	IF fbStopTx.bSettled THEN
		fbHourAngle.StopAxis := FALSE;
		fbDeclination.StopAxis := FALSE;
		_StopTelescope := FALSE;
	END_IF
END_IF
END_METHOD

METHOD PRIVATE _TrackTelescope : BOOL
VAR_INPUT
END_VAR
// send Dome position
THIS^.fbDome.Position := fAzimuthCurrent;
// Declination (including offest and pointing model)
fbDeclination.Position := fDeclinationApparent + fDeclinationOffset + fDeclinationPointingOffset;
// HourAngle
// change to -180 to 180 degree in HA
IF MODABS(fHourAngleApparent + F_HourAngleOffsetOnAxis(fHourAngleOffset, fDeclinationApparent)+ fHourAnglePointingOffset, 360) > 180 THEN
	fbHourAngle.Position := MODABS(fHourAngleApparent + F_HourAngleOffsetOnAxis(fHourAngleOffset, fDeclinationApparent)+ fHourAnglePointingOffset,360) - 360.0;
ELSE
	fbHourAngle.Position := MODABS(fHourAngleApparent + F_HourAngleOffsetOnAxis(fHourAngleOffset, fDeclinationApparent)+ fHourAnglePointingOffset,360);
END_IF


IF NOT fbHourAngle.Tracking THEN
	fbHourAngle.Velocity := 1.0;
	fbHourAngle.MoveAxis := TRUE;
	IF NOT fbHourAngle.Busy AND fbHourAngle.MoveDone THEN
		fbHourAngle.MoveAxis := FALSE;
		IF fbHourAngle.isTracking THEN
			fbHourAngle.Velocity := fHourAngleVelocity;
		END_IF
		fbHourAngle.Tracking := TRUE;
	END_IF
ELSE
	fbHourAngle.Velocity := fHourAngleVelocity;
END_IF


IF NOT fbDeclination.Tracking THEN
	fbDeclination.Velocity := 1.0;
	fbDeclination.MoveAxis := TRUE;
	IF NOT fbDeclination.Busy AND fbDeclination.MoveDone THEN
		fbDeclination.MoveAxis := FALSE;
		IF fbDeclination.isTracking THEN
			fbDeclination.Velocity := fDeclinationVelocity;
		END_IF
		fbDeclination.Tracking := TRUE;
	END_IF
ELSE
	fbDeclination.Velocity := fDeclinationVelocity;
END_IF
END_METHOD

PROPERTY AltAz : BROTLib.ST_AltAzCoordinate
GET
AltAz.Altitude 	:= fElevationCalc;
AltAz.Azimuth 	:= fAzimuthCalc;
END_GET
END_PROPERTY

{warning 'add property implementation'}
PROPERTY Altitude : LREAL
GET
Altitude := fElevationCurrent;
END_GET
END_PROPERTY

{warning 'add property implementation'}
PROPERTY Azimuth : LREAL
GET
Azimuth := fAzimuthCurrent;
END_GET
END_PROPERTY

PROPERTY CoverAutoOpen : BOOL
GET
CoverAutoOpen := bCoverAutoOpen;
END_GET
SET
bCoverAutoOpen := CoverAutoOpen;
END_SET
END_PROPERTY

{warning 'add property implementation'}
PROPERTY Declination : LREAL
GET
END_GET
END_PROPERTY

PROPERTY DeclinationOffset : LREAL
GET
DeclinationOffset := fDeclinationOffset;
END_GET
SET
fDeclinationOffset := DeclinationOffset;
END_SET
END_PROPERTY

//FB_Init is always available implicitly and it is used primarily for initialization.
//The return value is not evaluated. For a specific influence, you can also declare the
//methods explicitly and provide additional code there with the standard initialization
//code. You can evaluate the return value.
METHOD FB_Init: BOOL
VAR_INPUT
    bInitRetains	: BOOL; // TRUE: the retain variables are initialized (reset warm / reset cold)
    bInCopyCode		: BOOL;  // TRUE: the instance will be copied to the copy code afterward (online change)
	comm			: I_Comm;
END_VAR
THIS^.fbComm 				:= comm;
END_METHOD

METHOD Home : BOOL
bGoHomeChecked := TRUE;
// decide first (a home while not ready, powering on or parked is rejected, no longer waited for 2 min); a rejection writes nothing
IF NOT _AcceptMove(E_TCSCommand.gohome, E_TCSCommand.no_command) THEN
	RETURN;
END_IF
bHomeByCommand := TRUE;
bGoHomeActive := TRUE;
Home := TRUE;
END_METHOD

PROPERTY HourAngleOffset : LREAL
GET
HourAngleOffset := fHourAngleOffset;
END_GET
SET
fHourAngleOffset := HourAngleOffset;
END_SET
END_PROPERTY

METHOD Init : BOOL
bPowerChecked := TRUE;
// park wins in both orders and a stop is not overridden by a power-on (MONETcommon#87); this comes before AcceptInit, a pending
// park clears Initialized, so AcceptInit would accept. The in-place park (bSafeParked, up to 120 s) is refused as well.
IF bStopActive OR bParkActive OR bParkAfterStop OR bSafeParked THEN
    nInitRefusedCount := nInitRefusedCount + 1;
    bInitRefused := TRUE;
    IF bStopActive THEN
        sInitRefusedReason := 'stop in progress';
    ELSIF bSafeParked THEN
        sInitRefusedReason := 'in-place park in progress, ends within 120 s';
    ELSE
        sInitRefusedReason := 'park in progress, send stop to cancel it';
    END_IF
// AcceptInit refuses while a startup runs or completed (also across a transient interlock, -2).
ELSIF fbStartup.AcceptInit() THEN
    // nothing stale after the power-on starts: a pending move or home from before would run into it (park is kept, it is the safe direction)
    bGoHomeActive := FALSE;
    bGotoActive := FALSE;
    bSlewActive := FALSE;
    bTrackActive := FALSE;
    bPowerActive := TRUE;
    fReadyState := 0.7;
    // #159: an automatic stop leaves the sweep hold set with the axes enabled; a new power-on releases it
    fbHourAngle.bReleaseHold := TRUE;
    fbDeclination.bReleaseHold := TRUE;
END_IF
Init := TRUE;
END_METHOD

PROPERTY RaDec : BROTLib.ST_RaDecCoordinate
GET
RaDec.RightAscension	:= fRightAscensionCalc;
RaDec.Declination		:= fDeclinationCalc;
END_GET
END_PROPERTY

METHOD Reset : BOOL
bResetChecked := TRUE;
bResetRequest := TRUE;
END_METHOD

// READY_STATE as published on TELESCOPE.READY_STATE; BROTLib.FB_Comm_MQTT_Influx accepts the focus command only at 1 (BROTLib#74)
PROPERTY ReadyState : LREAL
GET
ReadyState := fReadyState;
END_GET
END_PROPERTY

{warning 'add property implementation'}
PROPERTY RightAscension : LREAL
GET
END_GET
END_PROPERTY

METHOD SetAltitudeOffset : BOOL
VAR_INPUT
	Offset	: LREAL;
END_VAR
END_METHOD

METHOD SetAzimuthOffset : BOOL
VAR_INPUT
	Offset	: LREAL;
END_VAR
END_METHOD

METHOD SetDeclinationOffset : BOOL
VAR_INPUT
	Offset	: LREAL;
END_VAR
fDeclinationOffset := Offset;
END_METHOD

METHOD SetDerotatorOffset : BOOL
VAR_INPUT
	Offset	: LREAL;
END_VAR
END_METHOD

METHOD SetRightAscensionOffset : BOOL
VAR_INPUT
	Offset	: LREAL;
END_VAR
fHourAngleOffset := -1.0*Offset;
END_METHOD

{warning 'add method implementation '}
METHOD Slew : BOOL
VAR_INPUT
	fAzimuth	: LREAL;
	fAltitude	: LREAL;
END_VAR
// #100: not while the telescope is not ready (parked, powering on, error). The request used to stay latched and
// fired unnoticed after the next power-on; a client sends init first and waits for ready.
bSlewChecked := TRUE;
// decided at arrival (F_CommandAcceptance): a rejected slew writes nothing, not even the target, and is never left pending
IF NOT _AcceptMove(E_TCSCommand.slew, E_TCSCommand.no_command) THEN
	RETURN;
END_IF
THIS^.fElevation 	:= fAltitude;
THIS^.fAzimuth 	:= fAzimuth;
bSlewActive		:= TRUE;
END_METHOD

METHOD Stop : BOOL
bStopChecked := TRUE;
// a stop ends a park that is queued behind a running stop (MONETcommon#213)
bParkAfterStop := FALSE;
// a repeated stop while a stop is running sends a new stop only to axes that are moving again and are not stopping already
// (BROTLib.FB_StopTransaction.Restart); the focus is stopped again as well (MONETcommon#96/#122)
IF bStopActive THEN
	_SetStopTxInputs();
	fbStopTx.Restart();
	IF fbFocus <> 0 THEN
		fbFocus.Stop();
	END_IF
END_IF
bStopActive := TRUE;
// MONETcommon#122: an explicit stop also stops a running focus move and holds the position reached; the automatic
// stops of the mount (horizon, pole zone) leave the focus alone
IF fbFocus <> 0 THEN
	fbFocus.Stop();
END_IF
END_METHOD

{warning 'add method implementation '}
METHOD Track : BOOL
VAR_INPUT
	fRightAscension	: LREAL;
	fDeclination	: LREAL;
END_VAR
// #100: see Slew(); a track request while the telescope is not ready is refused, not latched
bGotoChecked := TRUE;
bTrackChecked := TRUE;	// D4 (template body step S1.f): Track() and a bTrack edge in one scan are one command, as in MONETcommon
IF NOT _AcceptMove(E_TCSCommand.goto, E_TCSCommand.no_command) THEN
	RETURN;
END_IF
THIS^.fRightAscension	:= fRightAscension;
THIS^.fDeclination	:= fDeclination;
bGotoActive			:= TRUE;
END_METHOD

END_FUNCTION_BLOCK

(* stored: Version 1.1.0.1, ProductVersion 3.1.4024.15
   POU FB_TelescopeControl: Id {10c2c294-efcf-424f-afd3-75ac57a5e8bc}, SpecialFunc None
   Folder command methods: Id {f8e9235d-f769-45dd-a5d6-c3922581f371}
   Folder internal methods: Id {43f8a5dc-2166-4fdb-b436-34a8f62ea04a}
   Method _ScanBegin: Id {69ccb1e4-5ed8-4b33-8b32-527be9b9a8f0}
   Method _ReadInputs: Id {af4314b2-e999-4026-9f11-f74b6e7dc8b9}
   Method _ReadErrors: Id {98a12957-2fbf-495b-a37b-adfd985f2c64}
   Method _ErrorReaction: Id {c1780515-8c28-492e-9250-ace6f3e56191}
   Method _OnMoveEdgeAccepted: Id {ce98ff0a-3b98-4ad7-9bc7-3f0e8c90757d}
   Method _ApplyError: Id {79a0423b-d992-41a9-8dd9-6759ec5302b9}
   Method _ComputeTargets: Id {39a07f06-7eab-4842-b1ba-c5b3cddcad64}
   Method _Guards: Id {7de697b9-8dd1-4334-b9e3-11896fbb6ded}
   Method _Timers: Id {f5ac4a19-815a-48ce-aa91-a7e245e3fd2b}
   Method _RestartMoveTimeout: Id {a360d10e-6a59-40fc-8d4b-a2d75946ccc3}
   Method _ParkRequests: Id {844845fc-6fdb-4187-acd2-d29c542ffad9}
   Method _ParkPreStep: Id {05a3a385-eeb5-443f-91a3-5109b3bc5761}
   Method _EmergencyPark: Id {1fce47db-52d5-4e8f-8830-dce2ed613a3e}
   Method _AtRest: Id {02f74f7a-9e33-433b-bca7-1cc87c427b13}
   Method _InterruptPower: Id {b823f462-7c7e-4769-abb2-a73d057f39e5}
   Method _InterruptPark: Id {3a689de4-5be6-4fd3-8413-ed7b0cb662e7}
   Method _InterruptGoto: Id {b9c192ce-d0e0-4af4-8db8-6acabdc788c4}
   Method _InterruptSlew: Id {8aacbfb5-0cec-48bb-bf7c-31f98866be61}
   Method _InterruptGoHome: Id {79b6b6a9-c37f-4e8f-bc64-84e66edf7204}
   Method _AfterArbiter: Id {dda4d906-4b1f-4b0f-9b5d-ea64e8e7972f}
   Method _DropAxisCommands: Id {79f0235a-66ef-4f2e-a214-67cdf13e3e0b}
   Method _OnCommandChanged: Id {f346392c-2817-43c8-8907-287d92fd8956}
   Method _PowerOnStage: Id {7d1c9b36-52a4-4e0f-9c6d-3b8a41f0e5a2}
   Method _DoPowerOn: Id {454c13ff-2a44-40fe-9a9f-2af34564ef90}
   Method _DoPark: Id {b5264596-9ee8-4f0a-afa0-d22e2a0b4f11}
   Method _DoGoHome: Id {3b936219-2cea-4274-b961-23091a26a747}
   Method _DoGoto: Id {004b73df-348a-4a65-9a02-c72ce9d78c0f}
   Method _DoSlew: Id {4a88c6d3-4e35-43d1-93cd-57728314805b}
   Method _DoTrack: Id {b1bdd141-25f6-40a8-9621-d21903e5c547}
   Method _DoStop: Id {d21af247-3e6e-4829-b3e2-c95f07ff097e}
   Method _CommandTimeout: Id {338bbb57-390b-4e28-9d6e-df29401b077c}
   Method _AfterDispatch: Id {30cc36e7-894f-477a-80da-c4ca526c5b90}
   Method _UpdateStatus: Id {9a359329-5c54-4b0b-92c4-a82608059586}
   Method _ReadyStateParking: Id {88028a50-c2ca-4b03-acbc-fb2e926b6d1b}
   Method _IsSlewing: Id {2af0092a-3810-4785-ae7e-21e90e06e14d}
   Method _StopSettled: Id {ba012c82-2fb0-46d9-b276-40ac40c40998}
   Method _OnAbortStopReleased: Id {5e7ee996-2062-4ffc-b9db-4a9110b8e543}
   Method _ReleaseReset: Id {16858d95-be95-42c6-89a2-6f193b9ba85a}
   Method _SafeStateEndOfScan: Id {23aaa3a3-d319-45d1-a1a9-1948dea8722a}
   Method _TelemetryPeriod: Id {41c0c6f9-cff0-44ee-b857-7a38ef9d173e}
   Method _SendTelemetry: Id {c13d6275-e349-4a1b-a971-89e069fd0198}
   Method _EndOfScan: Id {abdb2eda-d02c-4cb5-b472-dab166d7ca3c}
   Folder properties: Id {65c2c08a-67b2-43de-bf16-65ce2beac397}
   Method _LogEvents: Id {2e11d121-0e66-42d3-bda8-e55c8ad61884}
   Method _CommandState: Id {dcfc70aa-b99e-45a8-9b01-d3cbca8d7345}
   Method _AcceptMove: Id {51edef40-3393-4d6a-a494-75062c704f44}
   Method _NoteRejected: Id {ccf0eb00-1bf6-40a0-b632-603d24022ec2}
   Method _AutoStop: Id {6f0d3a5e-2b91-4c78-8e14-7a9c5d3b1e02}
   Method _ParkInPlace: Id {8325b836-3a90-4df9-8d4a-8b6c11a8e16d}
   Method _HandleReset: Id {d3bbfeba-2cbb-4111-9ae3-4525c9154e5c}
   Method _ReadAxes: Id {fbf95db5-70d7-4355-ad80-f4cd75187122}
   Method _GotoTelescope: Id {43ebaf76-c0fc-41db-8c98-2f7671dc6b31}
   Method _HomeTelescope: Id {b2d9dfb4-bf7c-4f17-8ac5-7f074d6808c9}
   Method _ParkTelescope: Id {94a12771-4c75-4743-9ad3-850f66878f1f}
   Method _ResetErroredAxes: Id {5e8a3c17-9b42-4d06-a1f3-6c0d7e92b4a8}
   Method _PowerOnBlockedReason: Id {7c1e4b52-3a9d-4f60-b8e5-5d2f0a6c91e3}
   Method _PowerOn: Id {1dafa267-4251-4a45-a8e2-ae0ece289894}
   Method _SendTelemetryEquitorial: Id {2e72b74c-93b9-406f-985e-048a1bd902d8}
   Method _SlewTelescope: Id {4aaca2e7-2dba-4c2d-80b3-cd4dcc5ad38b}
   Method _SetStopTxInputs: Id {7c1b2e44-5d0a-4f63-9a1e-3b8d2f6c9e01}
   Method _StopTelescope: Id {cc9583d1-2578-4480-8aee-f6d55f373bf1}
   Method _TrackTelescope: Id {0dd53d55-2f74-4268-9438-8bb832d1c59b}
   Property AltAz: Id {82dbc2ee-80ef-40a3-8c1f-856f0af6c171}
   Get Get: Id {8533a901-9986-4274-8ee4-831d970f2e24}
   Property Altitude: Id {77878183-ff56-458d-9713-573db093fec2}
   Get Get: Id {d42084e4-5702-4d63-9998-7aed13913cd3}
   Property Azimuth: Id {af0c56f8-138d-4c6a-9afa-2054c20456bc}
   Get Get: Id {9755fb63-911d-4e5f-a9b2-82e25bd608d3}
   Property CoverAutoOpen: Id {a2921602-d837-46a8-9f8b-557b1c36a495}
   Get Get: Id {fbaf95b6-2065-4dce-8fd3-38db611cec44}
   Set Set: Id {7da2257e-bd6b-42e4-905b-2009b459922d}
   Property Declination: Id {9fcba06b-96da-4b28-85d9-479fe50b914c}
   Get Get: Id {6f7da282-4cc8-4a40-b385-90b0f4ce4349}
   Property DeclinationOffset: Id {653ff89d-921b-48cd-89fc-23fb937bb1d4}
   Get Get: Id {354ef6de-7ef9-4e01-82b0-872878ba7d1c}
   Set Set: Id {e59e1fb5-c6b1-429a-a0d7-2bdcae218f85}
   Method FB_Init: Id {034c34d9-521a-4d54-9624-e4d1bdeb670c}
   Method Home: Id {1ffeeb7f-e086-4ec6-b333-bf9ff24723c8}
   Property HourAngleOffset: Id {ac27a626-cead-47ea-868b-f24be3bdcddc}
   Get Get: Id {84bac731-b27e-41a5-ad78-15f19c3b02c7}
   Set Set: Id {7568e91e-7602-412a-ac33-275760080a3c}
   Method Init: Id {a631cabc-b5f9-4584-b7df-b1ee9d39f6ec}
   Property RaDec: Id {03d00136-4b42-4017-a768-650b9915ac54}
   Get Get: Id {51953765-9c9c-4236-b443-cc2f78a3c091}
   Method Reset: Id {f3acfef0-ab57-4326-aaf5-f5730beeec6a}
   Property ReadyState: Id {e6813a30-c227-4a62-a1fe-92138ff55729}
   Get Get: Id {4b91fc1d-55a3-4123-8f16-1d45dde7ec9c}
   Property RightAscension: Id {fbe599ea-0c8f-4d80-a746-e4e19f11c40d}
   Get Get: Id {db4c8087-9b17-4688-a0aa-8aab9120b914}
   Method SetAltitudeOffset: Id {25d1cab5-c5af-446c-a8a4-81112d093153}
   Method SetAzimuthOffset: Id {4fec041c-6825-4034-99a8-88dde866e4e2}
   Method SetDeclinationOffset: Id {f9c99137-b576-45ed-a746-cd632ae8760e}
   Method SetDerotatorOffset: Id {8c2a0fde-b71d-4d4a-9c60-3a9072f29e99}
   Method SetRightAscensionOffset: Id {10a7c758-0667-41d2-90bb-38e90ad006bf}
   Method Slew: Id {ba7a2a47-75f1-41c1-b2bd-a1c9f655c1f4}
   Method Stop: Id {e66d844d-991d-4af1-8b55-fe6740342385}
   Method Track: Id {6d7c3b1b-06e1-4002-b952-698198812e9b} *)
